// TIA Portal V21 export
// export: Created 2026-10-23T20:42:16.4522959Z, ExportSetting WithDefaults, DisplayName Totally Integrated Automation Portal, DisplayVersion V21 Update 1, DisplayName SINAMICS Startdrive Advanced, DisplayVersion V21 HF2, DisplayName SINAMICS Startdrive G110M, G120, G120C, G120D, G120P, G115D, DisplayVersion V21 HF2, DisplayName SINAMICS Startdrive G130, G150, S120, S150, G200, G220, S200, S210, S220, Innomotics MVD, DisplayVersion V21 HF2, DisplayName STEP 7 Professional, DisplayVersion V21 Update 1, DisplayName STEP 7 Safety, DisplayVersion V21, DisplayName Tech WebApplication, DisplayVersion V21, DisplayName WinCC Basic/Comfort/Advanced, DisplayVersion V21 Update 1, DisplayName WinCC Unified, DisplayVersion V21 Update 1
FUNCTION_BLOCK "F_FB_MainSafety"   // FB3, F_LAD
{ S7_Optimized_Access := 'TRUE' }
VERSION : 0.1
// stored: AutoNumber true, IsIECCheckEnabled false, UDAEnableTagReadback false
   VAR
      Enable : Bool;   // Schutztür geschlossen und Not-Halt in Ordnung / Guard closed and emergency stop ok
      Released : Bool;   // Maschine freigegeben / Machine released
      LogicRelease : Bool;   // Freigabe aus F_FC_Logic / Release from F_FC_Logic
   END_VAR
BEGIN

REGION Network 1: F-DB lesen / Read the F-DB
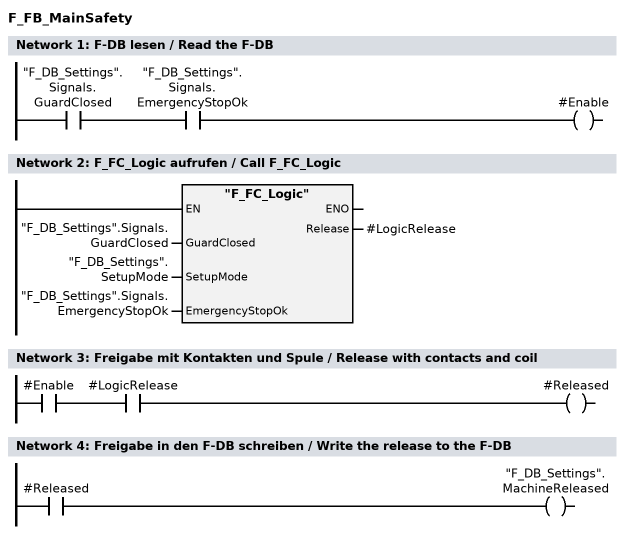
   RUNG wire#powerrail
      Contact( "F_DB_Settings".Signals.GuardClosed )
      Contact( "F_DB_Settings".Signals.EmergencyStopOk )
      Coil( #Enable )
   END_RUNG
   // the same network as SCL:
   #Enable := "F_DB_Settings".Signals.GuardClosed AND "F_DB_Settings".Signals.EmergencyStopOk;
END_REGION

REGION Network 2: F_FC_Logic aufrufen / Call F_FC_Logic
   RUNG wire#powerrail
      "F_FC_Logic"(GuardClosed := "F_DB_Settings".Signals.GuardClosed, SetupMode := "F_DB_Settings".SetupMode, EmergencyStopOk := "F_DB_Settings".Signals.EmergencyStopOk, Release => #LogicRelease)
   END_RUNG
   // the same network as SCL:
   "F_FC_Logic"(GuardClosed := "F_DB_Settings".Signals.GuardClosed,
                SetupMode := "F_DB_Settings".SetupMode,
                EmergencyStopOk := "F_DB_Settings".Signals.EmergencyStopOk,
                Release => #LogicRelease);
END_REGION

REGION Network 3: Freigabe mit Kontakten und Spule / Release with contacts and coil
   RUNG wire#powerrail
      Contact( #Enable )
      Contact( #LogicRelease )
      Coil( #Released )
   END_RUNG
   // the same network as SCL:
   #Released := #Enable AND #LogicRelease;
END_REGION

REGION Network 4: Freigabe in den F-DB schreiben / Write the release to the F-DB
   RUNG wire#powerrail
      Contact( #Released )
      Coil( "F_DB_Settings".MachineReleased )
   END_RUNG
   // the same network as SCL:
   "F_DB_Settings".MachineReleased := #Released;
END_REGION
END_FUNCTION_BLOCK
